Staubli VAL3: addlog.pgx

public program addlog(string x_sLog, num x_nType)
begin
  sLog[nIndex]=x_sLog
  nLogType[nIndex]=x_nType
  nIndex=(nIndex+1)%size(sLog)

end
